(* IEC 61131-3 sources: avi-aoi-management/scripts/ai-eval/ngau-nhien/kho/st-tv1-chong-doi/khung/src, 1 file *)

(* ---- ChongDoi.st ---- *)
FUNCTION_BLOCK ChongDoi
VAR_INPUT
    IN : BOOL;
    T_BAT : TIME;
    T_TAT : TIME;
END_VAR
VAR_OUTPUT
    Q : BOOL;
END_VAR
    (* TODO: cài đặt theo đề bài, dùng TON *)
    Q := FALSE;
END_FUNCTION_BLOCK
